Fanuc KAREL source: KT00915.KL

PROGRAM KT00915
%NOLOCKGROUP
VAR
  R1: REAL
  R2: REAL
  OUT: INTEGER
BEGIN
  R1 = 2.0
  R2 = 3.0
  R1 = 2.0
  R2 = 3.0
  OUT = STR_LEN(R1)
END KT00915
